SUBAPPLICATION Dauerfunktion (* Subapplication Type *)
  (* Standard: 61499-2 *)
  (* Version 1.0, 2023-01-29, Franz *)
  IMPORT DefaultPool::SoftKey_Licht;
  IMPORT isobus::UT::io::Softkey::SoftKeyActivationCode::SK_RELEASED;
  IMPORT DefaultPool::AuxInput_Licht;
  IMPORT isobus::UT::io::Auxiliary::IN::AuxiliaryState::AuxDisabled;
  IMPORT logiBUS::io::DQ::logiBUS_DO::Output_Q8;
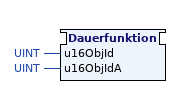
  VAR_INPUT
    u16ObjId : UINT;
    u16ObjIdA : UINT;
  END_VAR
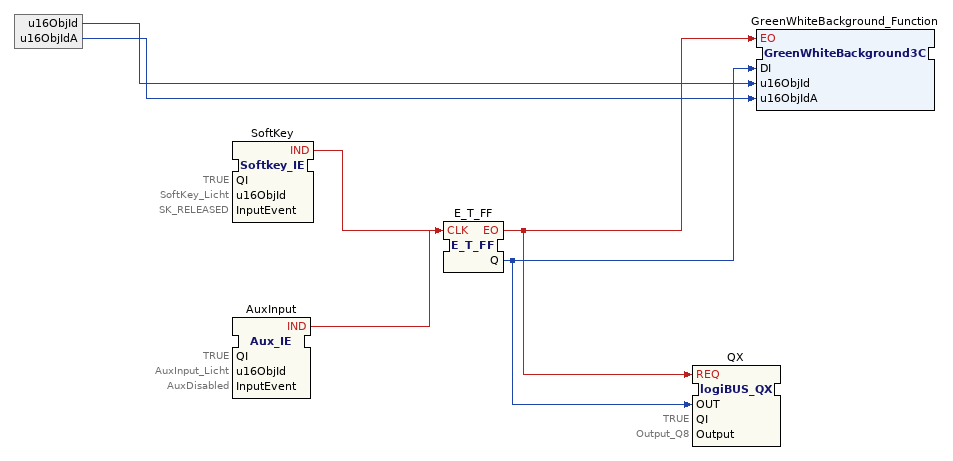
  FBS
    E_T_FF : iec61499::events::E_T_FF;
    QX : logiBUS::io::DQ::logiBUS_QX(QI := TRUE, Output := Output_Q8);
    SoftKey : isobus::UT::io::Softkey::Softkey_IE(QI := TRUE, u16ObjId := SoftKey_Licht, InputEvent := SK_RELEASED);
    AuxInput : isobus::UT::io::Auxiliary::IN::Aux_IE(QI := TRUE, u16ObjId := AuxInput_Licht, InputEvent := AuxDisabled);
  END_FBS
  SUBAPPS
    GreenWhiteBackground_Function : MyLib::sys::GreenWhiteBackground3C;
  END_SUBAPPS
  EVENT_CONNECTIONS
    E_T_FF.EO TO QX.REQ;
    E_T_FF.EO TO GreenWhiteBackground_Function.EO;
    SoftKey.IND TO E_T_FF.CLK;
    AuxInput.IND TO E_T_FF.CLK;
  END_CONNECTIONS
  DATA_CONNECTIONS
    E_T_FF.Q TO QX.OUT;
    E_T_FF.Q TO GreenWhiteBackground_Function.DI;
    u16ObjId TO GreenWhiteBackground_Function.u16ObjId;
    u16ObjIdA TO GreenWhiteBackground_Function.u16ObjIdA;
  END_CONNECTIONS
END_SUBAPPLICATION
